// #83: why F_CommandAcceptance rejected a command.
{attribute 'qualified_only'}
{attribute 'strict'}
TYPE E_CommandRejectReason :
(
	none := 0,
	estop,
	error,
	clock_invalid,
	stopping,
	powering_on,
	parking,
	parked,
	not_ready,
	gohome_active,
	init_required	// appended: MONETcommon#72 (a suspended telescope needs a new Init); only ever appended, the HMI reads it by value
);
END_TYPE

(* stored: Version 1.1.0.1, ProductVersion 3.1.4024.15
   DUT E_CommandRejectReason: Id {3e8d0ef8-4405-4709-be4f-fced965fe872} *)
